TEXTLIST TextList_TriBlenderUsage
  0 = 'Not in Use'
  1 = 'Marinada T1'
  2 = 'Marinada T2'
  3 = 'Marinada Stanbdy'
  4 = 'Color T3'
  5 = 'Color T4'
  6 = 'Color Standby'
   = ''
END_TEXTLIST

(* stored: Version 1.1.0.1, ProductVersion 3.1.4024.12
   TextList TextList_TriBlenderUsage: Id {959fde22-27f7-48e4-8947-2813d30f98b9} *)
